(* IEC 61131-3 sources: plc-hackathon-2026/hmi-me/generated, 1 file *)

(* ---- Team_Visu.st ---- *)
// HMI-only state and simulated-time chart axes. No control-strategy logic.
VAR_GLOBAL
 xResetArmed : BOOL;
 iAlarmPage : INT;
END_VAR
VAR_GLOBAL CONSTANT
 aHours : ARRAY[0..95] OF REAL := [-23.75, -23.50, -23.25, -23.00, -22.75, -22.50, -22.25, -22.00, -21.75, -21.50, -21.25, -21.00, -20.75, -20.50, -20.25, -20.00, -19.75, -19.50, -19.25, -19.00, -18.75, -18.50, -18.25, -18.00, -17.75, -17.50, -17.25, -17.00, -16.75, -16.50, -16.25, -16.00, -15.75, -15.50, -15.25, -15.00, -14.75, -14.50, -14.25, -14.00, -13.75, -13.50, -13.25, -13.00, -12.75, -12.50, -12.25, -12.00, -11.75, -11.50, -11.25, -11.00, -10.75, -10.50, -10.25, -10.00, -9.75, -9.50, -9.25, -9.00, -8.75, -8.50, -8.25, -8.00, -7.75, -7.50, -7.25, -7.00, -6.75, -6.50, -6.25, -6.00, -5.75, -5.50, -5.25, -5.00, -4.75, -4.50, -4.25, -4.00, -3.75, -3.50, -3.25, -3.00, -2.75, -2.50, -2.25, -2.00, -1.75, -1.50, -1.25, -1.00, -0.75, -0.50, -0.25, 0.00];
 aMonths : ARRAY[1..12] OF REAL := [1.0, 2.0, 3.0, 4.0, 5.0, 6.0, 7.0, 8.0, 9.0, 10.0, 11.0, 12.0];
END_VAR
